(* IEC 61131-3 sources: Summary-ETFA22/ahorn/test/benchmark/dissertation/PPU/ST (part 5) *)

        //End of: edu.kit.iti.formal.automation.st.IntroduceStateEnumVariable

        //Running pipeline step: edu.kit.iti.formal.automation.st.TranslationSfcToStOld$IntroduceTransitVariable

        //End of: edu.kit.iti.formal.automation.st.TranslationSfcToStOld$IntroduceTransitVariable

        //Running pipeline step: edu.kit.iti.formal.automation.st.TranslationSfcToStOld$TheBigStateCase

        CASE _state OF
            STATES_STAMP#Init:
                __transit := FALSE;
                IF TRUE THEN
                    __transit := TRUE;
                    _state := STATES_STAMP#Start_Stamp;
                END_IF

            STATES_STAMP#Start_Stamp:
                __transit := FALSE;
                Start_Stamp_active();
                IF interconnectStampStartCommand THEN
                    __transit := TRUE;
                    _state := STATES_STAMP#Green_Lamp;
                END_IF

            STATES_STAMP#Green_Lamp:
                __transit := FALSE;
                Green_Lamp_active();
                IF TRUE THEN
                    __transit := TRUE;
                    _state := STATES_STAMP#Stamp_Init_1;
                END_IF

            STATES_STAMP#Stamp_Init_1:
                __transit := FALSE;
                Stamp_Init_1_active();
                IF StampSliderSensorMovedIn THEN
                    __transit := TRUE;
                    _state := STATES_STAMP#Stamp_Init_2;
                END_IF

            STATES_STAMP#Stamp_Init_2:
                __transit := FALSE;
                Stamp_Init_2_active();
                IF StampSliderSensorMovedOut THEN
                    __transit := TRUE;
                    _state := STATES_STAMP#Stamp_Init_3;
                END_IF

            STATES_STAMP#Stamp_Init_3:
                __transit := FALSE;
                Stamp_Init_3_active();
                IF StampLowered THEN
                    __transit := TRUE;
                    _state := STATES_STAMP#Stamp_Init_4;
                END_IF

            STATES_STAMP#Stamp_Init_4:
                __transit := FALSE;
                Stamp_Init_4_active();
                IF StampUp THEN
                    __transit := TRUE;
                    _state := STATES_STAMP#Interstep;
                END_IF

            STATES_STAMP#Interstep:
                __transit := FALSE;
                Interstep_active();
                IF StartVar THEN
                    __transit := TRUE;
                    _state := STATES_STAMP#Intertsep_2;
                END_IF

            STATES_STAMP#Intertsep_2:
                __transit := FALSE;
                IF StampSliderFilled THEN
                    __transit := TRUE;
                    _state := STATES_STAMP#Step0;
                END_IF

            STATES_STAMP#Step0:
                __transit := FALSE;
                IF CraneUp THEN
                    __transit := TRUE;
                    _state := STATES_STAMP#StampSliderBack;
                END_IF

            STATES_STAMP#StampSliderBack:
                __transit := FALSE;
                StampSliderBack_active();
                IF StampSliderSensorMovedIn THEN
                    __transit := TRUE;
                    _state := STATES_STAMP#StampProcess;
                END_IF

            STATES_STAMP#StampProcess:
                __transit := FALSE;
                StampProcess_active();
                IF StampLowered THEN
                    __transit := TRUE;
                    _state := STATES_STAMP#Step1;
                END_IF

            STATES_STAMP#Step1:
                __transit := FALSE;
                Step1_active();
                IF interconnect THEN
                    __transit := TRUE;
                    _state := STATES_STAMP#StampSliderForward;
                END_IF

            STATES_STAMP#StampSliderForward:
                __transit := FALSE;
                StampSliderForward_active();
                IF StampSliderMovedOut THEN
                    __transit := TRUE;
                    _state := STATES_STAMP#Step2;
                END_IF

            STATES_STAMP#Step2:
                __transit := FALSE;
                IF (((AnalogCranePosition > 16160) AND (AnalogCranePosition < 16260)) AND NOT StampSliderFilled) THEN
                    __transit := TRUE;
                    _state := STATES_STAMP#Interstep;
                END_IF

                    END_CASE
        //End of: edu.kit.iti.formal.automation.st.TranslationSfcToStOld$TheBigStateCase

        //Running pipeline step: edu.kit.iti.formal.automation.st.SfcFlagIntroduction

    END_IF
    //End of: edu.kit.iti.formal.automation.st.SfcFlagIntroduction

END_FUNCTION_BLOCK

PROGRAM Main
    VAR_OUTPUT
        Actuator_AnalogCranePressure : INT := INT#0;
        Actuator_CraneLower : BOOL := FALSE;
        Actuator_CraneTurnClockwise : BOOL := FALSE;
        Actuator_CraneTurnCounterclockwise : BOOL := FALSE;
        Actuator_MagazinGreenLamp : BOOL := FALSE;
        Actuator_MagazinSlider : BOOL := FALSE;
        Actuator_MagazinVacuumOff : BOOL := FALSE;
        Actuator_MagazinVacuumOn : BOOL := FALSE;
        Actuator_MagazinWhiteLamp : BOOL := FALSE;
        Actuator_PusherY1 : BOOL := FALSE;
        Actuator_PusherY2 : BOOL := FALSE;
        Actuator_SorterConveyorTowardsCrane : BOOL := FALSE;
        Actuator_SorterConveyorTowardsStacker : BOOL := FALSE;
        Actuator_SorterGreenLampConveyor : BOOL := FALSE;
        Actuator_SorterWhiteLampConveyor : BOOL := FALSE;
        Actuator_StampGreenLamp : BOOL := FALSE;
        Actuator_StampPusher : BOOL := FALSE;
        Actuator_StampSliderMovedIn : BOOL := FALSE;
        Actuator_StampSliderMovedOut : BOOL := FALSE;
        Actuator_StampWhiteLamp : BOOL := FALSE;
    END_VAR

    VAR
        Conveyor : Conveyor := (SFCReset:=FALSE, Timer_Conveyor_Runtime:=(Q:=FALSE, PT:=UINT#0, IN:=FALSE, ET:=UINT#0), SorterStartButton:=FALSE, interconnect_Conveyor_Test:=FALSE, SorterConveyorTowardsCrane:=FALSE, interconnectConveyorStartCommand:=FALSE, SFCInit:=FALSE, interconnectConveyorTerminationCommand:=FALSE, SorterConveyorTowardsStacker:=FALSE, interconnect_Conveyor_Runtime:=FALSE, Timer_Conveyor_Test:=(Q:=FALSE, PT:=UINT#0, IN:=FALSE, ET:=UINT#0), SorterLightbarrierCraneInterface:=FALSE, SorterSwitchManuellAutomatic:=FALSE, StartVar:=FALSE, SorterGreenLampConveyor:=FALSE, StartCommandConveyor:=FALSE, Duration_Conveyor_Test:=TIME#1000.0ms, Duration_Conveyor_Runtime:=TIME#4500.0ms, SorterWhiteLampConveyor:=FALSE);
        Crane : Crane := (SliderMovedOut:=FALSE, CraneTurnCounterclockwise:=FALSE, WorkpieceReady:=FALSE, StampLowered:=FALSE, Duration1:=TIME#1500.0ms, StampSliderSensorMovedOut:=FALSE, TimeDelay_Timer_interconnect:=FALSE, MagazinOpticalSensor:=FALSE, StartVar:=FALSE, StartButtonMagazin:=FALSE, actualtime1:=TIME#, AnalogCranePressure:=INT#0, SFCReset:=FALSE, AnalogCranePosition:=INT#0, MagazinVacuumOff:=FALSE, CraneSucked:=FALSE, MagazinSlider:=FALSE, MagazinVacuumOn:=FALSE, interconnectCraneStartCommand:=FALSE, SFCInit:=FALSE, StartCommandCrane:=FALSE, TimeDelay_Timer_Duration:=TIME#50.0ms, interconnect:=FALSE, StampSliderFilled:=FALSE, CraneTurnClockwise:=FALSE, CraneUp:=FALSE, MagazinCapacitiveSensor:=FALSE, CraneLower:=FALSE, SliderNotMovedOut:=FALSE, CraneDown:=FALSE, TimeDelay_Timer:=(Q:=FALSE, PT:=UINT#0, IN:=FALSE, ET:=UINT#0), Timer1:=(Q:=FALSE, PT:=UINT#0, IN:=FALSE, ET:=UINT#0));
        Mag : Magazin := (SliderMovedOut:=FALSE, MagazinGreenLamp:=FALSE, interconnectMagazinStartCommand:=FALSE, SFCReset:=FALSE, AnalogCranePosition:=INT#0, CraneTurnCounterclockwise:=FALSE, MagazinVacuumOff:=FALSE, WorkpieceReady:=FALSE, CraneSucked:=FALSE, MagazinSlider:=FALSE, MagazinVacuumOn:=FALSE, MagazinWhiteLamp:=FALSE, SFCInit:=FALSE, StartCommandMagazin:=FALSE, CraneOnConveyor:=FALSE, CraneTurnClockwise:=FALSE, CraneUp:=FALSE, StartVar:=FALSE, CraneLower:=FALSE, SliderNotMovedOut:=FALSE, StartButtonMagazin:=FALSE, CraneOnMagazin:=FALSE, CraneDown:=FALSE);
        Pusher : Pusher := (Slide2_metal:=INT#1, Timer_Slide2_White:=(Q:=FALSE, PT:=UINT#0, IN:=FALSE, ET:=UINT#0), SorterPusher1MovedIn:=FALSE, SorterPusher2MovedIn:=FALSE, Slide3_white:=INT#1, Slide3_black:=INT#1, Timer_Slide1_Black:=(Q:=FALSE, PT:=UINT#0, IN:=FALSE, ET:=UINT#0), PusherY2:=FALSE, Priority_Var_Metal:=INT#3, PusherY1:=FALSE, SFCReset:=FALSE, SorterCapacitiveSensorPusher2:=FALSE, SorterCapacitiveSensorPusher1:=FALSE, Timer_Slide1_White:=(Q:=FALSE, PT:=UINT#0, IN:=FALSE, ET:=UINT#0), Timer_Slide2_Metal:=(Q:=FALSE, PT:=UINT#0, IN:=FALSE, ET:=UINT#0), Slide3_metal:=INT#1, Duration_Slide1_Metal:=TIME#300.0ms, Duration_Slide1_Black:=TIME#950.0ms, interconnect_Slide1_White:=FALSE, interconnect_Slide2_Metal:=FALSE, SorterPusher2MovedOut:=FALSE, Slide2_white:=INT#1, Priority_Var_Black:=INT#3, Duration_Slide2_Black:=TIME#2000.0ms, SorterLightnessSensorPusher2:=FALSE, SorterPusher1MovedOut:=FALSE, SorterStartButton:=FALSE, SorterLightnessSensorPusher1:=FALSE, Duration3:=TIME#200.0ms, Duration2:=TIME#2000.0ms, Slide1_black:=INT#1, interconnect_Slide2_White:=FALSE, SorterLightbarrierCraneInterface:=FALSE, StartVar:=FALSE, Duration_Slide2_White:=TIME#370.0ms, interconnect_Slide2_Black:=FALSE, SorterLightnessSensorPusher3:=FALSE, Slide1_white:=INT#1, interconnect3:=FALSE, interconnect2:=FALSE, interconnect_Slide1_Metal:=FALSE, Slide1_metal:=INT#1, SFCInit:=FALSE, Priority_Var_White:=INT#3, Slide2_black:=INT#1, Duration_Slide2_Metal:=TIME#370.0ms, interconnect_Slide1_Black:=FALSE, SorterLightnesssensorCraneInterfaceInverse:=FALSE, Timer_Slide1_Metal:=(Q:=FALSE, PT:=UINT#0, IN:=FALSE, ET:=UINT#0), Timer2:=(Q:=FALSE, PT:=UINT#0, IN:=FALSE, ET:=UINT#0), Timer_Slide2_Black:=(Q:=FALSE, PT:=UINT#0, IN:=FALSE, ET:=UINT#0), Duration_Slide1_White:=TIME#300.0ms, Timer3:=(Q:=FALSE, PT:=UINT#0, IN:=FALSE, ET:=UINT#0));
        Stamp : Stamp := (StampLowered:=FALSE, StampSliderSensorMovedOut:=FALSE, interconnectStampStartCommand:=FALSE, CraneOnConveyor:=FALSE, CranePositionStamp:=FALSE, StampSliderMovedOut:=FALSE, StartVar:=FALSE, StampPusher:=FALSE, StampWhiteLamp:=FALSE, StampPressure:=FALSE, SFCReset:=FALSE, StampGreenLamp:=FALSE, AnalogCranePosition:=INT#0, CraneSucked:=FALSE, Duration:=TIME#500.0ms, SFCInit:=FALSE, StampStartButton:=FALSE, StampSliderSensorMovedIn:=FALSE, interconnect:=FALSE, StampSliderFilled:=FALSE, CraneUp:=FALSE, StampSliderMovedIn:=FALSE, Timer:=(Q:=FALSE, PT:=UINT#0, IN:=FALSE, ET:=UINT#0), StartCommandStamp:=FALSE, CraneDown:=FALSE, StampUp:=FALSE);
    END_VAR

    VAR_INPUT
        Sensor_AnalogCranePosition : INT := INT#0;
        Sensor_CraneDown : BOOL := FALSE;
        Sensor_CraneOnConveyor : BOOL := FALSE;
        Sensor_CraneOnMagazin : BOOL := FALSE;
        Sensor_CranePosition : BOOL := FALSE;
        Sensor_CranePositionStamp : BOOL := FALSE;
        Sensor_CraneSucked : BOOL := FALSE;
        Sensor_CraneUp : BOOL := FALSE;
        Sensor_MagazinCapacitiveSensor : BOOL := FALSE;
        Sensor_MagazinEmergencyStop : BOOL := FALSE;
        Sensor_MagazinOpticalSensor : BOOL := FALSE;
        Sensor_MagazinSwitchManuellAutomatic : BOOL := FALSE;
        Sensor_SliderMovedOut : BOOL := FALSE;
        Sensor_SliderNotMovedOut : BOOL := FALSE;
        Sensor_SorterCapacitiveSensorPusher1 : BOOL := FALSE;
        Sensor_SorterCapacitiveSensorPusher2 : BOOL := FALSE;
        Sensor_SorterEmergencyStop : BOOL := FALSE;
        Sensor_SorterLightbarrierCraneInterface : BOOL := FALSE;
        Sensor_SorterLightnessSensorPusher1 : BOOL := FALSE;
        Sensor_SorterLightnessSensorPusher2 : BOOL := FALSE;
        Sensor_SorterLightnessSensorPusher3 : BOOL := FALSE;
        Sensor_SorterLightnesssensorCraneInterfaceInverse : BOOL := FALSE;
        Sensor_SorterPusher1MovedIn : BOOL := FALSE;
        Sensor_SorterPusher1MovedOut : BOOL := FALSE;
        Sensor_SorterPusher2MovedIn : BOOL := FALSE;
        Sensor_SorterPusher2MovedOut : BOOL := FALSE;
        Sensor_SorterStartButton : BOOL := FALSE;
        Sensor_SorterSwitchManuellAutomatic : BOOL := FALSE;
        Sensor_StampEmergencyStop : BOOL := FALSE;
        Sensor_StampLowered : BOOL := FALSE;
        Sensor_StampSliderFilled : BOOL := FALSE;
        Sensor_StampSliderSensorMovedIn : BOOL := FALSE;
        Sensor_StampSliderSensorMovedOut : BOOL := FALSE;
        Sensor_StampStartButton : BOOL := FALSE;
        Sensor_StampSwitchManuellAutomatic : BOOL := FALSE;
        Sensor_StampUp : BOOL := FALSE;
        Sensor_StartButtonMagazin : BOOL := FALSE;
        Sensor_WorkpieceReady : BOOL := FALSE;
    END_VAR

    Mag.SliderNotMovedOut := Sensor_SliderNotMovedOut;
    Mag.SliderMovedOut := Sensor_SliderMovedOut;
    Mag.CraneOnMagazin := Sensor_CraneOnMagazin;
    Mag.CraneDown := Sensor_CraneDown;
    Mag.CraneUp := Sensor_CraneUp;
    Mag.CraneOnConveyor := Sensor_CraneOnConveyor;
    Mag.WorkpieceReady := Sensor_WorkpieceReady;
    Mag.AnalogCranePosition := Sensor_AnalogCranePosition;
    Mag.StartButtonMagazin := Sensor_StartButtonMagazin;
    Actuator_MagazinSlider := Mag.MagazinSlider;
    Actuator_MagazinGreenLamp := Mag.MagazinGreenLamp;
    Crane.CraneUp := Sensor_CraneUp;
    Crane.CraneDown := Sensor_CraneDown;
    Crane.CraneSucked := Sensor_CraneSucked;
    Crane.MagazinCapacitiveSensor := Sensor_MagazinCapacitiveSensor;
    Crane.SliderMovedOut := Sensor_SliderMovedOut;
    Crane.WorkpieceReady := Sensor_WorkpieceReady;
    Crane.MagazinOpticalSensor := Sensor_MagazinOpticalSensor;
    Crane.StampSliderFilled := Sensor_StampSliderFilled;
    Crane.StampSliderSensorMovedOut := Sensor_StampSliderSensorMovedOut;
    Crane.StampLowered := Sensor_StampLowered;
    Crane.AnalogCranePosition := Sensor_AnalogCranePosition;
    Crane.StartButtonMagazin := Sensor_StartButtonMagazin;
    Actuator_CraneTurnCounterclockwise := Crane.CraneTurnCounterclockwise;
    Actuator_CraneTurnClockwise := Crane.CraneTurnClockwise;
    Actuator_CraneLower := Crane.CraneLower;
    Actuator_MagazinVacuumOff := Crane.MagazinVacuumOff;
    Actuator_MagazinVacuumOn := Crane.MagazinVacuumOn;
    Actuator_AnalogCranePressure := Crane.AnalogCranePressure;
    Stamp.StampSliderSensorMovedOut := Sensor_StampSliderSensorMovedOut;
    Stamp.StampSliderSensorMovedIn := Sensor_StampSliderSensorMovedIn;
    Stamp.StampSliderFilled := Sensor_StampSliderFilled;
    Stamp.StampUp := Sensor_StampUp;
    Stamp.StampLowered := Sensor_StampLowered;
    Stamp.CraneDown := Sensor_CraneDown;
    Stamp.CraneUp := Sensor_CraneUp;
    Stamp.CraneSucked := Sensor_CraneSucked;
    Stamp.CranePositionStamp := Sensor_CranePositionStamp;
    Stamp.CraneOnConveyor := Sensor_CraneOnConveyor;
    Stamp.AnalogCranePosition := Sensor_AnalogCranePosition;
    Stamp.StampStartButton := Sensor_StampStartButton;
    Actuator_StampSliderMovedOut := Stamp.StampSliderMovedOut;
    Actuator_StampSliderMovedIn := Stamp.StampSliderMovedIn;
    Actuator_StampWhiteLamp := Stamp.StampWhiteLamp;
    Actuator_StampPusher := Stamp.StampPusher;
    Actuator_StampGreenLamp := Stamp.StampGreenLamp;
    Conveyor.SorterStartButton := Sensor_SorterStartButton;
    Conveyor.SorterSwitchManuellAutomatic := Sensor_SorterSwitchManuellAutomatic;
    Conveyor.SorterLightbarrierCraneInterface := Sensor_SorterLightbarrierCraneInterface;
    Actuator_SorterConveyorTowardsStacker := Conveyor.SorterConveyorTowardsStacker;
    Actuator_SorterConveyorTowardsCrane := Conveyor.SorterConveyorTowardsCrane;
    Actuator_SorterGreenLampConveyor := Conveyor.SorterGreenLampConveyor;
    Actuator_SorterWhiteLampConveyor := Conveyor.SorterWhiteLampConveyor;
    Pusher.SorterLightnesssensorCraneInterfaceInverse := Sensor_SorterLightnesssensorCraneInterfaceInverse;
    Pusher.SorterLightbarrierCraneInterface := Sensor_SorterLightbarrierCraneInterface;
    Pusher.SorterCapacitiveSensorPusher1 := Sensor_SorterCapacitiveSensorPusher1;
    Pusher.SorterLightnessSensorPusher1 := Sensor_SorterLightnessSensorPusher1;
    Pusher.SorterCapacitiveSensorPusher2 := Sensor_SorterCapacitiveSensorPusher2;
    Pusher.SorterLightnessSensorPusher2 := Sensor_SorterLightnessSensorPusher2;
    Pusher.SorterLightnessSensorPusher3 := Sensor_SorterLightnessSensorPusher3;
    Pusher.SorterPusher1MovedOut := Sensor_SorterPusher1MovedOut;
    Pusher.SorterPusher1MovedIn := Sensor_SorterPusher1MovedIn;
    Pusher.SorterPusher2MovedOut := Sensor_SorterPusher2MovedOut;
    Pusher.SorterPusher2MovedIn := Sensor_SorterPusher2MovedIn;
    Pusher.SorterStartButton := Sensor_SorterStartButton;
    Actuator_PusherY1 := Pusher.PusherY1;
    Actuator_PusherY2 := Pusher.PusherY2;
    IF ((Sensor_SorterEmergencyStop AND Sensor_StampEmergencyStop) AND Sensor_MagazinEmergencyStop) THEN
        Mag();
        Crane();
        Stamp();
        Conveyor();
        Pusher();
        IF ((Actuator_SorterGreenLampConveyor AND Actuator_MagazinGreenLamp) AND Actuator_StampGreenLamp) THEN
            IF (((Stamp.StartCommandStamp AND Crane.StartCommandCrane) AND Conveyor.StartCommandConveyor) AND Mag.StartCommandMagazin) THEN
                Crane.StartVar := TRUE;
                Conveyor.StartVar := TRUE;
                Mag.StartVar := TRUE;
                Pusher.StartVar := TRUE;
                Stamp.StartVar := TRUE;
            END_IF
        END_IF
        Crane.SFCReset := FALSE;
        Conveyor.SFCReset := FALSE;
        Mag.SFCReset := FALSE;
        Pusher.SFCReset := FALSE;
        Stamp.SFCReset := FALSE;
    ELSIF ((NOT Sensor_SorterEmergencyStop OR NOT Sensor_StampEmergencyStop) OR NOT Sensor_MagazinEmergencyStop) THEN
        Actuator_MagazinSlider := FALSE;
        Actuator_CraneLower := FALSE;
        Actuator_MagazinVacuumOn := FALSE;
        Actuator_MagazinVacuumOff := TRUE;
        Actuator_MagazinGreenLamp := FALSE;
        Actuator_CraneTurnCounterclockwise := FALSE;
        Actuator_CraneTurnClockwise := FALSE;
        Actuator_SorterConveyorTowardsStacker := FALSE;
        Actuator_SorterConveyorTowardsCrane := FALSE;
        Actuator_SorterGreenLampConveyor := FALSE;
        Actuator_PusherY1 := FALSE;
        Actuator_PusherY2 := FALSE;
        Actuator_StampSliderMovedOut := TRUE;
        Actuator_StampSliderMovedIn := FALSE;
        Actuator_StampGreenLamp := FALSE;
        Actuator_StampPusher := FALSE;
        Actuator_AnalogCranePressure := INT#0;
        Crane.SFCReset := TRUE;
        Conveyor.SFCReset := TRUE;
        Mag.SFCReset := TRUE;
        Pusher.SFCReset := TRUE;
        Stamp.SFCReset := TRUE;
        Crane.StartVar := FALSE;
        Conveyor.StartVar := FALSE;
        Mag.StartVar := FALSE;
        Pusher.StartVar := FALSE;
        Stamp.StartVar := FALSE;
    END_IF
END_PROGRAM
FUNCTION_BLOCK CTD

    VAR_INPUT
        CD : BOOL := FALSE;
        LD : BOOL := FALSE;
        PV : INT := INT#0;
    END_VAR

    VAR_OUTPUT
        CV : INT := INT#0;
        Q : BOOL := FALSE;
    END_VAR

    IF LD THEN
        CV := PV;
    ELSIF (CU AND (CV > INT#0)) THEN
        CV := (CV - INT#1);
    END_IF
    Q := (CV <= INT#0);
END_FUNCTION_BLOCK

FUNCTION_BLOCK CTU

    VAR_INPUT
        CU : BOOL := FALSE;
        PV : INT := INT#0;
        R : BOOL := FALSE;
    END_VAR

    VAR_OUTPUT
        CV : INT := INT#0;
        Q : BOOL := FALSE;
    END_VAR

    IF R THEN
        CV := INT#0;
    ELSIF (CU AND (CV < PV)) THEN
        CV := (CV + INT#1);
    END_IF
    Q := (CV >= PV);
END_FUNCTION_BLOCK

FUNCTION_BLOCK R_TRIG

    VAR_INPUT
        CLK : BOOL := FALSE;
    END_VAR

    VAR
        M : BOOL := FALSE;
    END_VAR

    VAR_OUTPUT
        Q : BOOL := FALSE;
    END_VAR

    Q := (CLK AND NOT M);
    M := CLK;
END_FUNCTION_BLOCK

FUNCTION_BLOCK F_TRIG

    VAR_INPUT
        CLK : BOOL := FALSE;
    END_VAR

    VAR
        M : BOOL := TRUE;
    END_VAR

    VAR_OUTPUT
        Q : BOOL := FALSE;
    END_VAR

    Q := (NOT CLK AND NOT M);
    M := NOT CLK;
END_FUNCTION_BLOCK

FUNCTION SEL : ANY

    VAR_INPUT
        G : BOOL := FALSE;
        a : ANY;
        b : ANY;
    END_VAR

    VAR_OUTPUT
        SEL : ANY;
    END_VAR

    IF G THEN
        SEL := a;
    ELSE
        SEL := b;
    END_IF
END_FUNCTION

FUNCTION MAX : ANY_INT

    VAR_OUTPUT
        MAX : ANY_INT;
    END_VAR

    VAR_INPUT
        in0 : ANY_INT;
        in1 : ANY_INT;
    END_VAR

    MAX := sel((in0 >= in1), in0, in1);
END_FUNCTION

FUNCTION MIN : ANY_INT

    VAR_OUTPUT
        MIN : ANY_INT;
    END_VAR

    VAR_INPUT
        in0 : ANY_INT;
        in1 : ANY_INT;
    END_VAR

    MIN := sel((in0 <= in1), in0, in1);
END_FUNCTION

FUNCTION LIMIT : INT

    VAR_OUTPUT
        LIMIT : INT := INT#0;
    END_VAR

    VAR_INPUT
        in : ANY_INT;
        max : ANY_INT;
        min : ANY_INT;
    END_VAR

    LIMIT := MAX(min, MIN(in, max));
END_FUNCTION

FUNCTION ERROR : ANY

    VAR_OUTPUT
        ERROR : ANY;
    END_VAR

    VAR
        msg : STRING := WSTRING#"";
    END_VAR

END_FUNCTION

FUNCTION SMV : ANY

    VAR_OUTPUT
        SMV : ANY;
    END_VAR

    VAR_INPUT
        code : STRING := WSTRING#"";
    END_VAR

END_FUNCTION

FUNCTION_BLOCK TON

    VAR_OUTPUT
        ET : UINT := UINT#0;
        Q : BOOL := FALSE;
    END_VAR

    VAR_INPUT
        IN : BOOL := FALSE;
        PT : UINT := UINT#0;
    END_VAR

    IF IN THEN
        Q := (ET = UINT#0);
        IF (ET > UINT#0) THEN
            ET := (ET - UINT#1);
        ELSE
            ET := UINT#0;
        END_IF
    ELSE
        Q := FALSE;
        ET := PT;
    END_IF
END_FUNCTION_BLOCK

TYPE SFC_STEPS: STRUCT

        T :TIME
        X :BOOL
        _T :TIME
        _X :BOOLEND_STRUCT;

END_TYPE

TYPE
    STATES_CONVEYOR : (Init, Start_Conveyor, Green_Lamp, Conveyor_Init, Conveyor_init_2, Interstep, Step0, Conveyor_Towards_Stacker, Runtime_Conveyor, Conveyor_pause, Conveyor_Stop_Empty_Magazin);
    STATES_CRANE : (Init, Start_Crane, Crane_Init, Crane_Init_2, Interstep, Interstep_2, TimeDelay, Interstep_3, Turn_Right, Magazin_Stop, Crane_Lower, Step0, Crane_Lift_Magazin, Crane_Turn_Left_NOT_Metallic, Crane_On_Conveyor, Stamp_Pressure_Profile_Set_Metallic, Crane_Lift_Magazin_Metallic, Crane_Turn_Left_Metallic, Crane_On_Stamp_Metallic, release_Workpiece, Crane_Go_Up, Stamp_Pressure_Profile_Set_White, Crane_Lift_Magazin_White, Crane_Turn_Left_White, Crane_On_Stamp_White, release_Workpiece_White, Crane_Go_Up_White, Step3, Step2, pause, Turn_Right_Black, Magazin_Stop_Black, Crane_Lift_NOT_Metallic_Black, Crane_Turn_Left_NOT_Metallic_Black, Crane_On_Conveyor_Not_Metallica_Black, release_Black, Crane_Lift_Conveyor_Black, Crane_Turn_Left_Back_To_Stamp, Crane_On_Stamp_Stop_Black, Step4, Reset_interconnect, Lower_Crane, Suck_At_Stamp, Crane_Lift_At_Stamp, Crane_Turn_Left_From_Stamp, Crane_On_Conveyor_Metallic, release, Crane_Lift_Conveyor, No_Workpiece_ready, Crane_Turn_Left_Metallic2, Crane_On_Stamp_Metallic2, Interstep_4, Crane_On_Stamp_Metallic2_Lower, Suck_At_Stamp2, Crane_Lift_At_Stamp2, Crane_Turn_Right_From_Stamp, Crane_On_Conveyor_Metallic2, release2, Crane_Lift_Conveyor2, Turn_Right_Final, Magazin_Stop_Final);
    STATES_MAGAZIN : (Init, Start_Magazin, Green_Lamp, Magazin_Init, Magazin_Init_2, Interstep, convey, Step0, Slider_Move_Back, Step1);
    STATES_PUSHER : (Init, Interstep, Interstep_2, Check_For_Black, Third_Slide_black_workpieces, Wait_Black, Reset_interconnect3, Second_Slide_black_workpieces, Second_Slide_Timer_Black, PusherY2_Move_Out_Black, Wait_Y2_Black, PusherY2_Move_In_Black, Reset_interconnect_Slide2_Black, First_Slide_black_workpieces, First_Slide_Timer_Black, PusherY1_Move_Out_Black, Wait_Y1_Black, PusherY1_Move_In_Black, Reset_interconnect_Slide1_Black, Check_For_White, First_Slide_white_workpieces, First_Slide_Timer_White, PusherY1_Move_Out_White, Wait_Y1_White, PusherY1_Move_In_White, Reset_interconnect_Slide1_White, Second_Slide_white_workpieces, Second_Test_For_White, Second_Slide_Timer_White, PusherY2_Move_Out_White, Wait_Y2_White, PusherY2_Move_In_White, Reset_interconnect_Slide2_White, Third_Slide_white_workpieces, Wait_White, Reset_interconnect_Slide3_White, Check_For_Metal, First_Slide_metal_workpieces, First_Slide_Timer_Metal, PusherY1_Move_Out_Metal, Wait_Y1_Metal, PusherY1_Move_In_Metal, Reset_interconnect_Slide1_Metal, Second_Slide_metal_workpieces, Second_Test_For_Metal, Second_Slide_Timer_Metal, PusherY2_Move_Out_Metal, Wait_Y2_Metal, PusherY2_Move_In_Metal, Reset_interconnect_Slide2_Metal, Third_Slide_metal_workpieces, Wait_Metal, Reset_interconnect_Slide3_Metal);
    STATES_STAMP : (Init, Start_Stamp, Green_Lamp, Stamp_Init_1, Stamp_Init_2, Stamp_Init_3, Stamp_Init_4, Interstep, Intertsep_2, Step0, StampSliderBack, StampProcess, Step1, StampSliderForward, Step2);
END_TYPE

(* ---- Scenario1_Final.st ---- *)
TYPE
    CraneStates : (CraneSFCInit, StartCrane, CraneInit, CraneInit2, Interstep, Interstep2, TimeDelay, TurnRight,
                   InterstepCheckWorkpiece, StackStop, CraneLiftStack, CraneTurnLeft, CraneOnConveyorState,
                   release, CraneLiftConveyor, CraneStop);
    StackStates : (StackSFCInit, StartStack, GreenLamp, StackInit, StackInit2, Interstep, convey, Step0,
                   SliderMoveBack, Step1);
END_TYPE

FUNCTION_BLOCK Crane
VAR_INPUT
    CraneDown : BOOL := FALSE;
    CraneOnConveyor : BOOL := FALSE;
    CraneOnStack : BOOL := FALSE;
    CraneSucked : BOOL := FALSE;
    CraneUp : BOOL := FALSE;
    SFCReset : BOOL := FALSE;
    SliderMovedOut : BOOL := FALSE;
    SliderNotMovedOut : BOOL := FALSE;
    StartButtonStack : BOOL := FALSE;
    StartVar : BOOL := FALSE;
    WorkpieceReady : BOOL := FALSE;
END_VAR
VAR
    SFCInit : BOOL := FALSE;
    SFCPause : BOOL := FALSE;
    CraneState : CraneStates := CraneStates#CraneSFCInit;
    Timer : TON;
    TimerDuration : TIME := TIME#50.0ms;
    Timerinterconnect : BOOL := FALSE;
    interconnectCraneStartCommand : BOOL := FALSE;
END_VAR
VAR_OUTPUT
    CraneLower : BOOL := FALSE;
    CraneTurnClockwise : BOOL := FALSE;
    CraneTurnCounterClockwise : BOOL := FALSE;
    StackVacuumOff : BOOL := FALSE;
    StackVacuumOn : BOOL := FALSE;
    StartCommandCrane : BOOL := FALSE;
END_VAR

IF (SFCInit OR SFCReset) THEN
    CraneDown := FALSE;
    CraneLower := FALSE;
    CraneOnConveyor := FALSE;
    CraneOnStack := FALSE;
    CraneSucked := FALSE;
    CraneTurnClockwise := FALSE;
    CraneTurnCounterClockwise := FALSE;
    CraneUp := FALSE;
    StackVacuumOff := FALSE;
    StackVacuumOn := FALSE;
    SFCInit := FALSE;
    SFCReset := FALSE;
    SliderMovedOut := FALSE;
    SliderNotMovedOut := FALSE;
    StartButtonStack := FALSE;
    StartCommandCrane := FALSE;
    StartVar := FALSE;
    Timer.ET := INT#0;
    Timer.IN := FALSE;
    Timer.PT := INT#0;
    Timer.Q := FALSE;
    TimerDuration := TIME#50ms;
    Timerinterconnect := FALSE;
    WorkpieceReady := FALSE;
    CraneState := CraneStates#CraneSFCInit;
    interconnectCraneStartCommand := FALSE;
END_IF;

IF NOT (SFCInit OR SFCPause) THEN
    CASE CraneState OF
        CraneStates#CraneSFCInit:
            IF TRUE THEN
                CraneState := CraneStates#StartCrane;
            END_IF;

        CraneStates#StartCrane:
            CraneLower := FALSE;
            StackVacuumOff := TRUE;
            StackVacuumOn := FALSE;
            CraneTurnCounterClockwise := FALSE;
            CraneTurnClockwise := FALSE;
            StartVar := FALSE;
            StartCommandCrane := FALSE;
            IF (StartButtonStack = TRUE) THEN
                interconnectCraneStartCommand := TRUE;
            END_IF;
            IF interconnectCraneStartCommand THEN
                CraneState := CraneStates#CraneInit;
            END_IF;

        CraneStates#CraneInit:
            CraneLower := TRUE;
            interconnectCraneStartCommand := FALSE;
            IF CraneDown THEN
                CraneState := CraneStates#CraneInit2;
            END_IF;

        CraneStates#CraneInit2:
            CraneLower := FALSE;
            IF CraneUp THEN
                CraneState := CraneStates#Interstep;
            END_IF;

        CraneStates#Interstep:
            StartCommandCrane := TRUE;
            IF StartVar THEN
                CraneState := CraneStates#Interstep2;
            END_IF;

        CraneStates#Interstep2:
            IF SliderMovedOut THEN
                CraneState := CraneStates#TimeDelay;
            END_IF;

        CraneStates#TimeDelay:
            Timer(IN := TRUE, PT := TimerDuration);
            Timerinterconnect := Timer.Q;
            IF Timerinterconnect THEN
                CraneState := CraneStates#TurnRight;
            END_IF;

        CraneStates#TurnRight:
            CraneTurnClockwise := TRUE;
            CraneTurnCounterClockwise := FALSE;
            IF CraneOnStack THEN
                CraneState := CraneStates#InterstepCheckWorkpiece;
            END_IF;

        CraneStates#InterstepCheckWorkpiece:
            IF WorkpieceReady THEN
                CraneState := CraneStates#StackStop;
            ELSIF NOT WorkpieceReady THEN
                CraneState := CraneStates#CraneStop;
            END_IF;

        CraneStates#StackStop:
            CraneTurnClockwise := FALSE;
            CraneTurnCounterClockwise := FALSE;
            StackVacuumOn := TRUE;
            StackVacuumOff := FALSE;
            CraneLower := TRUE;
            IF CraneSucked THEN
                CraneState := CraneStates#CraneLiftStack;
            END_IF;

        CraneStates#CraneLiftStack:
            CraneLower := FALSE;
            IF CraneUp THEN
                CraneState := CraneStates#CraneTurnLeft;
            END_IF;

        CraneStates#CraneTurnLeft:
            CraneTurnCounterClockwise := TRUE;
            CraneTurnClockwise := FALSE;
            IF CraneOnConveyor THEN
                CraneState := CraneStates#CraneOnConveyorState;
            END_IF;

        CraneStates#CraneOnConveyorState:
            CraneTurnCounterClockwise := FALSE;
            CraneTurnClockwise := FALSE;
            CraneLower := TRUE;
            IF CraneDown THEN
                CraneState := CraneStates#release;
            END_IF;

        CraneStates#release:
            StackVacuumOff := TRUE;
            StackVacuumOn := FALSE;
            IF TRUE THEN
                CraneState := CraneStates#CraneLiftConveyor;
            END_IF;

        CraneStates#CraneLiftConveyor:
            CraneLower := FALSE;
            IF TRUE THEN
                CraneState := CraneStates#Interstep;
            END_IF;

        CraneStates#CraneStop:
            IF TRUE THEN
                CraneState := CraneStates#StartCrane;
            END_IF;
    END_CASE;
END_IF;
END_FUNCTION_BLOCK

FUNCTION_BLOCK Stack
VAR_INPUT
    CraneDown : BOOL := FALSE;
    CraneOnConveyor : BOOL := FALSE;
    CraneOnStack : BOOL := FALSE;
    CraneSucked : BOOL := FALSE;
    CraneUp : BOOL := FALSE;
    SFCReset : BOOL := FALSE;
    SliderMovedOut : BOOL := FALSE;
    SliderNotMovedOut : BOOL := FALSE;
    StartButtonStack : BOOL := FALSE;
    StartVar : BOOL := FALSE;
    WorkpieceReady : BOOL := FALSE;
END_VAR
VAR
    SFCInit : BOOL := FALSE;
    SFCPause : BOOL := FALSE;
    StackState : StackStates := StackStates#StackSFCInit;
    interconnectStackStartCommand : BOOL := FALSE;
END_VAR
VAR_OUTPUT
    StackGreenLamp : BOOL := FALSE;
    StackSlider : BOOL := FALSE;
    StartCommandStack : BOOL := FALSE;
END_VAR

IF (SFCInit OR SFCReset) THEN
    CraneDown := FALSE;
    CraneOnConveyor := FALSE;
    CraneOnStack := FALSE;
    CraneSucked := FALSE;
    CraneUp := FALSE;
    StackGreenLamp := FALSE;
    StackSlider := FALSE;
    SFCInit := FALSE;
    SFCReset := FALSE;
    SliderMovedOut := FALSE;
    SliderNotMovedOut := FALSE;
    StartButtonStack := FALSE;
    StartCommandStack := FALSE;
    StartVar := FALSE;
    WorkpieceReady := FALSE;
    StackState := StackStates#StackSFCInit;
    interconnectStackStartCommand := FALSE;
END_IF;

IF NOT (SFCInit OR SFCPause) THEN
    CASE StackState OF
        StackStates#StackSFCInit:
            IF TRUE THEN
                StackState := StackStates#StartStack;
            END_IF;

        StackStates#StartStack:
            StackSlider := FALSE;
            StackGreenLamp := FALSE;
            StartVar := FALSE;
            StartCommandStack := FALSE;
            IF (StartButtonStack = TRUE) THEN
                interconnectStackStartCommand := TRUE;
            END_IF;
            IF interconnectStackStartCommand THEN
                StackState := StackStates#GreenLamp;
            END_IF;

        StackStates#GreenLamp:
            StackGreenLamp := TRUE;
            interconnectStackStartCommand := FALSE;
            IF TRUE THEN
                StackState := StackStates#StackInit;
            END_IF;

        StackStates#StackInit:
            StackSlider := TRUE;
            IF TRUE THEN
                StackState := StackStates#StackInit2;
            END_IF;

        StackStates#StackInit2:
            StackSlider := FALSE;
            IF TRUE THEN
                StackState := StackStates#Interstep;
            END_IF;

        StackStates#Interstep:
            StartCommandStack := TRUE;
            IF StartVar THEN
                StackState := StackStates#convey;
            END_IF;

        StackStates#convey:
            IF SliderNotMovedOut THEN
                StackSlider := TRUE;
            END_IF;
            IF CraneOnStack THEN
                StackState := StackStates#Step0;
            END_IF;

        StackStates#Step0:
            IF CraneDown THEN
                StackState := StackStates#SliderMoveBack;
            END_IF;

        StackStates#SliderMoveBack:
            IF ((SliderMovedOut = TRUE) AND (SliderNotMovedOut = FALSE)) THEN
                StackSlider := FALSE;
            END_IF;
            IF CraneUp THEN
                StackState := StackStates#Step1;
            END_IF;

        StackStates#Step1:
            IF CraneOnConveyor THEN
                StackState := StackStates#Interstep;
            END_IF;
    END_CASE;
END_IF;
END_FUNCTION_BLOCK

PROGRAM Main
VAR_INPUT
    SensorCraneDown : BOOL := FALSE;
    SensorCraneOnConveyor : BOOL := FALSE;
    SensorCraneOnStack : BOOL := FALSE;
    SensorCranePosition : BOOL := FALSE;
    SensorCraneSucked : BOOL := FALSE;
    SensorCraneUp : BOOL := FALSE;
    SensorStackEmergencyStop : BOOL := FALSE;
    SensorStackSwitchManuellAutomatic : BOOL := FALSE;
    SensorSliderMovedOut : BOOL := FALSE;
    SensorSliderNotMovedOut : BOOL := FALSE;
    SensorStartButtonStack : BOOL := FALSE;
    SensorWorkpieceReady : BOOL := FALSE;
END_VAR
VAR
    Crane : Crane;
    Stack : Stack;
END_VAR
VAR_OUTPUT
    ActuatorCraneLower : BOOL := FALSE;
    ActuatorCraneTurnClockwise : BOOL := FALSE;
    ActuatorCraneTurnCounterClockwise : BOOL := FALSE;
    ActuatorStackGreenLamp : BOOL := FALSE;
    ActuatorStackSlider : BOOL := FALSE;
    ActuatorStackVacuumOff : BOOL := FALSE;
    ActuatorStackVacuumOn : BOOL := FALSE;
    ActuatorStackWhiteLamp : BOOL := FALSE;
END_VAR
Stack.SliderNotMovedOut := SensorSliderNotMovedOut;
Stack.SliderMovedOut := SensorSliderMovedOut;
Stack.CraneOnStack := SensorCraneOnStack;
Stack.CraneDown := SensorCraneDown;
Stack.CraneUp := SensorCraneUp;
Stack.CraneOnConveyor := SensorCraneOnConveyor;
Stack.WorkpieceReady := SensorWorkpieceReady;
Stack.StartButtonStack := SensorStartButtonStack;
ActuatorStackSlider := Stack.StackSlider;
ActuatorStackGreenLamp := Stack.StackGreenLamp;
Crane.WorkpieceReady := SensorWorkpieceReady;
Crane.CraneUp := SensorCraneUp;
Crane.CraneOnConveyor := SensorCraneOnConveyor;
Crane.CraneDown := SensorCraneDown;
Crane.CraneSucked := SensorCraneSucked;
Crane.CraneOnStack := SensorCraneOnStack;
Crane.SliderMovedOut := SensorSliderMovedOut;
Crane.StartButtonStack := SensorStartButtonStack;
ActuatorCraneTurnCounterClockwise := Crane.CraneTurnCounterClockwise;
ActuatorCraneTurnClockwise := Crane.CraneTurnClockwise;
ActuatorCraneLower := Crane.CraneLower;
ActuatorStackVacuumOff := Crane.StackVacuumOff;
ActuatorStackVacuumOn := Crane.StackVacuumOn;
IF SensorStackEmergencyStop THEN
    Stack();
    Crane();
    IF ActuatorStackGreenLamp THEN
        IF (Crane.StartCommandCrane AND Stack.StartCommandStack) THEN
            Crane.StartVar := TRUE;
            Stack.StartVar := TRUE;
        END_IF;
    END_IF;
    Crane.SFCReset := FALSE;
    Stack.SFCReset := FALSE;
ELSIF NOT SensorStackEmergencyStop THEN
    ActuatorStackSlider := FALSE;
    ActuatorCraneLower := FALSE;
    ActuatorStackVacuumOn := FALSE;
    ActuatorStackVacuumOff := TRUE;
    ActuatorStackGreenLamp := FALSE;
    ActuatorCraneTurnCounterClockwise := FALSE;
    ActuatorCraneTurnClockwise := FALSE;
    Crane.SFCReset := TRUE;
    Stack.SFCReset := TRUE;
    Crane.StartVar := FALSE;
    Stack.StartVar := FALSE;
END_IF;
END_PROGRAM

FUNCTION_BLOCK TON
VAR_INPUT
    IN : BOOL;
    PT : TIME;
END_VAR
VAR
    running : BOOL;
END_VAR
VAR_TEMP
    timeout : BOOL;
END_VAR
VAR_OUTPUT
    Q : BOOL;
    ET : TIME;
END_VAR
timeout := NONDETERMINISTIC_BOOL();
IF NOT IN THEN
    Q := FALSE;
    running := FALSE;
ELSIF NOT running AND NOT Q THEN
    running := TRUE;
ELSIF running AND NOT Q THEN
    Q := timeout;
    running := NOT Q;
END_IF;
ET := NONDETERMINISTIC_TIME();
END_FUNCTION_BLOCK

(* ---- Scenario2_Final.st ---- *)
TYPE
    CraneStates : (CraneSFCInit, StartCrane, CraneInit, CraneInit2, Interstep, Interstep2, TimeDelay, TurnRight,
                   InterstepCheckWorkpiece, StackStop, Step0, CraneLiftStack, CraneTurnLeftNOTMetallic,
                   CraneOnConveyorState, CraneLiftStackMetallic, CraneTurnLeftMetallic, CraneOnConveyorMetallic,
                   release, CraneLiftConveyor, CraneStop);
    StackStates : (StackSFCInit, StartStack, GreenLamp, StackInit, StackInit2, Interstep, convey, Step0, SliderMoveBack,
                   Step1);
END_TYPE

FUNCTION_BLOCK Crane
VAR_INPUT
    CraneDown : BOOL := FALSE;
    CraneOnConveyor : BOOL := FALSE;
    CraneOnStack : BOOL := FALSE;
    CraneSucked : BOOL := FALSE;
    CraneUp : BOOL := FALSE;
    StackCapacitiveSensor : BOOL := FALSE;
    SFCReset : BOOL := FALSE;
    SliderMovedOut : BOOL := FALSE;
    SliderNotMovedOut : BOOL := FALSE;
    StartButtonStack : BOOL := FALSE;
    StartVar : BOOL := FALSE;
    WorkpieceReady : BOOL := FALSE;
END_VAR
VAR
    SFCInit : BOOL := FALSE;
    SFCPause : BOOL := FALSE;
    CraneState : CraneStates := CraneStates#CraneSFCInit;
    Timer : TON;
    TimerDuration : TIME := TIME#50.0ms;
    Timerinterconnect : BOOL := FALSE;
    interconnectCraneStartCommand : BOOL := FALSE;
END_VAR
VAR_OUTPUT
    CraneLower : BOOL := FALSE;
    CraneTurnClockwise : BOOL := FALSE;
    CraneTurnCounterClockwise : BOOL := FALSE;
    StackVacuumOff : BOOL := FALSE;
    StackVacuumOn : BOOL := FALSE;
    StartCommandCrane : BOOL := FALSE;
END_VAR

IF (SFCInit OR SFCReset) THEN
    CraneDown := FALSE;
    CraneLower := FALSE;
    CraneOnConveyor := FALSE;
    CraneOnStack := FALSE;
    CraneSucked := FALSE;
    CraneTurnClockwise := FALSE;
    CraneTurnCounterClockwise := FALSE;
    CraneUp := FALSE;
    StackCapacitiveSensor := FALSE;
    StackVacuumOff := FALSE;
    StackVacuumOn := FALSE;
    SFCInit := FALSE;
    SFCReset := FALSE;
    SliderMovedOut := FALSE;
    SliderNotMovedOut := FALSE;
    StartButtonStack := FALSE;
    StartCommandCrane := FALSE;
    StartVar := FALSE;
    Timer.ET := INT#0;
    Timer.IN := FALSE;
    Timer.PT := INT#0;
    Timer.Q := FALSE;
    TimerDuration := TIME#50ms;
    Timerinterconnect := FALSE;
    WorkpieceReady := FALSE;
    CraneState := CraneStates#CraneSFCInit;
    interconnectCraneStartCommand := FALSE;
END_IF;

IF NOT (SFCInit OR SFCPause) THEN
    CASE CraneState OF
        CraneStates#CraneSFCInit:
            IF TRUE THEN
                CraneState := CraneStates#StartCrane;
            END_IF;

        CraneStates#StartCrane:
            CraneLower := FALSE;
            StackVacuumOff := TRUE;
            StackVacuumOn := FALSE;
            CraneTurnCounterClockwise := FALSE;
            CraneTurnClockwise := FALSE;
            StartVar := FALSE;
            StartCommandCrane := FALSE;
            IF (StartButtonStack = TRUE) THEN
                interconnectCraneStartCommand := TRUE;
            END_IF;
            IF interconnectCraneStartCommand THEN
                CraneState := CraneStates#CraneInit;
            END_IF;

        CraneStates#CraneInit:
            CraneLower := TRUE;
            interconnectCraneStartCommand := FALSE;
            IF CraneDown THEN
                CraneState := CraneStates#CraneInit2;
            END_IF;

        CraneStates#CraneInit2:
            CraneLower := FALSE;
            IF CraneUp THEN
                CraneState := CraneStates#Interstep;
            END_IF;

        CraneStates#Interstep:
            StartCommandCrane := TRUE;
            IF StartVar THEN
                CraneState := CraneStates#Interstep2;
            END_IF;

        CraneStates#Interstep2:
            IF SliderMovedOut THEN
                CraneState := CraneStates#TimeDelay;
            END_IF;

        CraneStates#TimeDelay:
            Timer(IN := TRUE, PT := TimerDuration);
            Timerinterconnect := Timer.Q;
            IF Timerinterconnect THEN
                CraneState := CraneStates#TurnRight;
            END_IF;

        CraneStates#TurnRight:
            CraneTurnClockwise := TRUE;
            CraneTurnCounterClockwise := FALSE;
            IF CraneOnStack THEN
                CraneState := CraneStates#InterstepCheckWorkpiece;
            END_IF;

        CraneStates#InterstepCheckWorkpiece:
            IF WorkpieceReady THEN
                CraneState := CraneStates#StackStop;
            ELSIF NOT WorkpieceReady THEN
                CraneState := CraneStates#CraneStop;
            END_IF;

        CraneStates#StackStop:
            CraneTurnClockwise := FALSE;
            CraneTurnCounterClockwise := FALSE;
            StackVacuumOn := TRUE;
            StackVacuumOff := FALSE;
            CraneLower := TRUE;
            IF CraneSucked THEN
                CraneState := CraneStates#Step0;
            END_IF;

        CraneStates#Step0:
            IF NOT StackCapacitiveSensor THEN
                CraneState := CraneStates#CraneLiftStack;
            ELSIF StackCapacitiveSensor THEN
                CraneState := CraneStates#CraneLiftStackMetallic;
            END_IF;

        CraneStates#CraneLiftStack:
            CraneLower := FALSE;
            IF CraneUp THEN
                CraneState := CraneStates#CraneTurnLeftNOTMetallic;
            END_IF;

        CraneStates#CraneTurnLeftNOTMetallic:
            CraneTurnCounterClockwise := TRUE;
            CraneTurnClockwise := FALSE;
            IF CraneOnConveyor THEN
                CraneState := CraneStates#CraneOnConveyorState;
            END_IF;

        CraneStates#CraneOnConveyorState:
            CraneTurnCounterClockwise := FALSE;
            CraneTurnClockwise := FALSE;
            CraneLower := TRUE;
            IF CraneDown THEN
                CraneState := CraneStates#release;
            END_IF;

        CraneStates#CraneLiftStackMetallic:
            CraneLower := FALSE;
            IF CraneUp THEN
                CraneState := CraneStates#CraneTurnLeftMetallic;
            END_IF;

        CraneStates#CraneTurnLeftMetallic:
            CraneTurnCounterClockwise := TRUE;
            CraneTurnClockwise := FALSE;
            IF CraneOnConveyor THEN
                CraneState := CraneStates#CraneOnConveyorMetallic;
            END_IF;

        CraneStates#CraneOnConveyorMetallic:
            CraneTurnCounterClockwise := FALSE;
            CraneTurnClockwise := FALSE;
            CraneLower := TRUE;
            IF CraneDown THEN
                CraneState := CraneStates#release;
            END_IF;

        CraneStates#release:
            StackVacuumOff := TRUE;
            StackVacuumOn := FALSE;
            IF TRUE THEN
                CraneState := CraneStates#CraneLiftConveyor;
            END_IF;

        CraneStates#CraneLiftConveyor:
            CraneLower := FALSE;
            IF TRUE THEN
                CraneState := CraneStates#Interstep;
            END_IF;

        CraneStates#CraneStop:
            IF TRUE THEN
                CraneState := CraneStates#StartCrane;
            END_IF;
    END_CASE;
END_IF;
END_FUNCTION_BLOCK

FUNCTION_BLOCK Stack
VAR_INPUT
    CraneDown : BOOL := FALSE;
    CraneOnConveyor : BOOL := FALSE;
    CraneOnStack : BOOL := FALSE;
    CraneSucked : BOOL := FALSE;
    CraneUp : BOOL := FALSE;
    SFCReset : BOOL := FALSE;
    SliderMovedOut : BOOL := FALSE;
    SliderNotMovedOut : BOOL := FALSE;
    StartButtonStack : BOOL := FALSE;
    StartVar : BOOL := FALSE;
    WorkpieceReady : BOOL := FALSE;
END_VAR
VAR
    SFCInit : BOOL := FALSE;
    SFCPause : BOOL := FALSE;
    StackState : StackStates := StackStates#StackSFCInit;
    interconnectStackStartCommand : BOOL := FALSE;
END_VAR
VAR_OUTPUT
    CraneLower : BOOL := FALSE;
    CraneTurnClockwise : BOOL := FALSE;
    CraneTurnCounterClockwise : BOOL := FALSE;
    StackGreenLamp : BOOL := FALSE;
    StackSlider : BOOL := FALSE;
    StackVacuumOff : BOOL := FALSE;
    StackVacuumOn : BOOL := FALSE;
    StackWhiteLamp : BOOL := FALSE;
    StartCommandStack : BOOL := FALSE;
END_VAR

IF (SFCInit OR SFCReset) THEN
    CraneDown := FALSE;
    CraneLower := FALSE;
    CraneOnConveyor := FALSE;
    CraneOnStack := FALSE;
    CraneSucked := FALSE;
    CraneTurnClockwise := FALSE;
    CraneTurnCounterClockwise := FALSE;
    CraneUp := FALSE;
    StackGreenLamp := FALSE;
    StackSlider := FALSE;
    StackVacuumOff := FALSE;
    StackVacuumOn := FALSE;
    StackWhiteLamp := FALSE;
    SFCInit := FALSE;
    SFCReset := FALSE;
    SliderMovedOut := FALSE;
    SliderNotMovedOut := FALSE;
    StartButtonStack := FALSE;
    StartCommandStack := FALSE;
    StartVar := FALSE;
    WorkpieceReady := FALSE;
    StackState := StackStates#StackSFCInit;
    interconnectStackStartCommand := FALSE;
END_IF;

IF NOT (SFCInit OR SFCPause) THEN
    CASE StackState OF
        StackStates#StackSFCInit:
            IF TRUE THEN
                StackState := StackStates#StartStack;
            END_IF;

        StackStates#StartStack:
            StackSlider := FALSE;
            StackGreenLamp := FALSE;
            StartVar := FALSE;
            StartCommandStack := FALSE;
            IF (StartButtonStack = TRUE) THEN
                interconnectStackStartCommand := TRUE;
            END_IF;
            IF interconnectStackStartCommand THEN
                StackState := StackStates#GreenLamp;
            END_IF;

        StackStates#GreenLamp:
            StackGreenLamp := TRUE;
            interconnectStackStartCommand := FALSE;
            IF TRUE THEN
                StackState := StackStates#StackInit;
            END_IF;

        StackStates#StackInit:
            StackSlider := TRUE;
            IF TRUE THEN
                StackState := StackStates#StackInit2;
            END_IF;

        StackStates#StackInit2:
            StackSlider := FALSE;
            IF TRUE THEN
                StackState := StackStates#Interstep;
            END_IF;

        StackStates#Interstep:
            StartCommandStack := TRUE;
            IF StartVar THEN
                StackState := StackStates#convey;
            END_IF;

        StackStates#convey:
            IF SliderNotMovedOut THEN
                StackSlider := TRUE;
            END_IF;
            IF CraneOnStack THEN
                StackState := StackStates#Step0;
            END_IF;

        StackStates#Step0:
            IF CraneDown THEN
                StackState := StackStates#SliderMoveBack;
            END_IF;

        StackStates#SliderMoveBack:
            IF ((SliderMovedOut = TRUE) AND (SliderNotMovedOut = FALSE)) THEN
                StackSlider := FALSE;
            END_IF;
            IF CraneUp THEN
                StackState := StackStates#Step1;
            END_IF;

        StackStates#Step1:
            IF CraneOnConveyor THEN
                StackState := StackStates#Interstep;
            END_IF;
    END_CASE;
END_IF;
END_FUNCTION_BLOCK

PROGRAM Main
VAR_INPUT
    SensorCraneDown : BOOL := FALSE;
    SensorCraneOnConveyor : BOOL := FALSE;
    SensorCraneOnStack : BOOL := FALSE;
    SensorCranePosition : BOOL := FALSE;
    SensorCranePositionStamp : BOOL := FALSE;
    SensorCraneSucked : BOOL := FALSE;
    SensorCraneUp : BOOL := FALSE;
    SensorStackCapacitiveSensor : BOOL := FALSE;
    SensorStackEmergencyStop : BOOL := FALSE;
    SensorStackOpticalSensor : BOOL := FALSE;
    SensorStackSwitchManuellAutomatic : BOOL := FALSE;
    SensorSliderMovedOut : BOOL := FALSE;
    SensorSliderNotMovedOut : BOOL := FALSE;
    SensorStartButtonStack : BOOL := FALSE;
    SensorWorkpieceReady : BOOL := FALSE;
END_VAR
VAR
    Crane : Crane;
    Stack : Stack;
END_VAR
VAR_OUTPUT
    ActuatorCraneLower : BOOL := FALSE;
    ActuatorCraneTurnClockwise : BOOL := FALSE;
    ActuatorCraneTurnCounterClockwise : BOOL := FALSE;
    ActuatorStackGreenLamp : BOOL := FALSE;
    ActuatorStackSlider : BOOL := FALSE;
    ActuatorStackVacuumOff : BOOL := FALSE;
    ActuatorStackVacuumOn : BOOL := FALSE;
    ActuatorStackWhiteLamp : BOOL := FALSE;
END_VAR
Stack.SliderNotMovedOut := SensorSliderNotMovedOut;
Stack.SliderMovedOut := SensorSliderMovedOut;
Stack.CraneOnStack := SensorCraneOnStack;
Stack.CraneDown := SensorCraneDown;
Stack.CraneUp := SensorCraneUp;
Stack.CraneOnConveyor := SensorCraneOnConveyor;
Stack.WorkpieceReady := SensorWorkpieceReady;
Stack.StartButtonStack := SensorStartButtonStack;
ActuatorStackSlider := Stack.StackSlider;
ActuatorStackGreenLamp := Stack.StackGreenLamp;
Crane.WorkpieceReady := SensorWorkpieceReady;
Crane.CraneUp := SensorCraneUp;
Crane.CraneOnConveyor := SensorCraneOnConveyor;
Crane.CraneDown := SensorCraneDown;
Crane.CraneSucked := SensorCraneSucked;
Crane.CraneOnStack := SensorCraneOnStack;
Crane.StackCapacitiveSensor := SensorStackCapacitiveSensor;
Crane.SliderMovedOut := SensorSliderMovedOut;
Crane.StartButtonStack := SensorStartButtonStack;
ActuatorCraneTurnCounterClockwise := Crane.CraneTurnCounterClockwise;
ActuatorCraneTurnClockwise := Crane.CraneTurnClockwise;
ActuatorCraneLower := Crane.CraneLower;
ActuatorStackVacuumOff := Crane.StackVacuumOff;
ActuatorStackVacuumOn := Crane.StackVacuumOn;
IF SensorStackEmergencyStop THEN
    Stack();
    Crane();
    IF ActuatorStackGreenLamp THEN
        IF (Crane.StartCommandCrane AND Stack.StartCommandStack) THEN
            Crane.StartVar := TRUE;
            Stack.StartVar := TRUE;
        END_IF;
    END_IF;
    Crane.SFCReset := FALSE;
    Stack.SFCReset := FALSE;
ELSIF NOT SensorStackEmergencyStop THEN
    ActuatorStackSlider := FALSE;
    ActuatorCraneLower := FALSE;
    ActuatorStackVacuumOn := FALSE;
    ActuatorStackVacuumOff := TRUE;
    ActuatorStackGreenLamp := FALSE;
    ActuatorCraneTurnCounterClockwise := FALSE;
    ActuatorCraneTurnClockwise := FALSE;
    Crane.SFCReset := TRUE;
    Stack.SFCReset := TRUE;
    Crane.StartVar := FALSE;
    Stack.StartVar := FALSE;
END_IF;
END_PROGRAM

FUNCTION_BLOCK TON
VAR_INPUT
    IN : BOOL;
    PT : TIME;
END_VAR
VAR
    running : BOOL;
END_VAR
VAR_TEMP
    timeout : BOOL;
END_VAR
VAR_OUTPUT
    Q : BOOL;
    ET : TIME;
END_VAR
timeout := NONDETERMINISTIC_BOOL();
IF NOT IN THEN
    Q := FALSE;
    running := FALSE;
ELSIF NOT running AND NOT Q THEN
    running := TRUE;
ELSIF running AND NOT Q THEN
    Q := timeout;
    running := NOT Q;
END_IF;
ET := NONDETERMINISTIC_TIME();
END_FUNCTION_BLOCK

(* ---- Scenario3_Final.st ---- *)
TYPE
    CraneStates : (CraneSFCInit, StartCrane, CraneInit, CraneInit2, Interstep, Interstep2, TimeDelay, TurnRight,
                   InterstepCheckWorkpiece, StackStop, Step0, CraneLiftStack, CraneTurnLeftNOTMetallic,
                   CraneOnConveyorState, CraneLiftStackMetallic, CraneTurnLeftMetallic, CraneOnStampMetallic,
                   releaseWorkpiece, CraneGoUp, pause, Resetinterconnect, LowerCrane, SuckAtStamp, CraneLiftAtStamp,
                   CraneTurnLeftFromStamp, CraneOnConveyorMetallic, release, CraneLiftConveyor, WaitAtStamp, Step2);
    StackStates : (StackSFCInit, StartStack, GreenLamp, StackInit, StackInit2, Interstep, convey, Step0, SliderMoveBack,
                   Step1);
    StampStates : (StampSFCInit, StartStamp, GreenLamp, StampInit1, StampInit2, StampInit3, StampInit4, Interstep,
                   Interstep2, Step0, StampSliderBack, StampProcess, Step1, StampSliderForward, Step2);
END_TYPE

FUNCTION_BLOCK Crane
VAR_INPUT
    CraneDown : BOOL := FALSE;
    CraneOnConveyor : BOOL := FALSE;
    CraneOnStack : BOOL := FALSE;
    CranePositionStamp : BOOL := FALSE;
    CraneSucked : BOOL := FALSE;
    CraneUp : BOOL := FALSE;
    StackCapacitiveSensor : BOOL := FALSE;
    SFCReset : BOOL := FALSE;
    SliderMovedOut : BOOL := FALSE;
    SliderNotMovedOut : BOOL := FALSE;
    StampLowered : BOOL := FALSE;
    StampSliderFilled : BOOL := FALSE;
    StartButtonStack : BOOL := FALSE;
    StartVar : BOOL := FALSE;
    WorkpieceReady : BOOL := FALSE;
END_VAR
VAR
    Duration1 : TIME := TIME#1500.0ms;
    SFCInit : BOOL := FALSE;
    SFCPause : BOOL := FALSE;
    CraneState : CraneStates := CraneStates#CraneSFCInit;
    Timer : TON;
    TimerDuration : TIME := TIME#50.0ms;
    Timerinterconnect : BOOL := FALSE;
    Timer1 : TON;
    interconnect : BOOL := FALSE;
    interconnectCraneStartCommand : BOOL := FALSE;
END_VAR
VAR_OUTPUT
    CraneLower : BOOL := FALSE;
    CraneTurnClockwise : BOOL := FALSE;
    CraneTurnCounterClockwise : BOOL := FALSE;
    StackVacuumOff : BOOL := FALSE;
    StackVacuumOn : BOOL := FALSE;
    StartCommandCrane : BOOL := FALSE;
END_VAR

IF (SFCInit OR SFCReset) THEN
    CraneDown := FALSE;
    CraneLower := FALSE;
    CraneOnConveyor := FALSE;
    CraneOnStack := FALSE;
    CranePositionStamp := FALSE;
    CraneSucked := FALSE;
    CraneTurnClockwise := FALSE;
    CraneTurnCounterClockwise := FALSE;
    CraneUp := FALSE;
    Duration1 := TIME#1500ms;
    StackCapacitiveSensor := FALSE;
    StackVacuumOff := FALSE;
    StackVacuumOn := FALSE;
    SFCInit := FALSE;
    SFCReset := FALSE;
    SliderMovedOut := FALSE;
    SliderNotMovedOut := FALSE;
    StampLowered := FALSE;
    StampSliderFilled := FALSE;
    StartButtonStack := FALSE;
    StartCommandCrane := FALSE;
    StartVar := FALSE;
    Timer.ET := INT#0;
    Timer.IN := FALSE;
    Timer.PT := INT#0;
    Timer.Q := FALSE;
    TimerDuration := TIME#50ms;
    Timerinterconnect := FALSE;
    Timer1.ET := INT#0;
    Timer1.IN := FALSE;
    Timer1.PT := INT#0;
    Timer1.Q := FALSE;
    WorkpieceReady := FALSE;
    CraneState := CraneStates#CraneSFCInit;
    interconnect := FALSE;
    interconnectCraneStartCommand := FALSE;
END_IF;

IF NOT (SFCInit OR SFCPause) THEN
    CASE CraneState OF
        CraneStates#CraneSFCInit:
            IF TRUE THEN
                CraneState := CraneStates#StartCrane;
            END_IF;

        CraneStates#StartCrane:
            CraneLower := FALSE;
            StackVacuumOff := TRUE;
            StackVacuumOn := FALSE;
            CraneTurnCounterClockwise := FALSE;
            CraneTurnClockwise := FALSE;
            StartVar := FALSE;
            StartCommandCrane := FALSE;
            IF (StartButtonStack = TRUE) THEN
                interconnectCraneStartCommand := TRUE;
            END_IF;
            IF interconnectCraneStartCommand THEN
                CraneState := CraneStates#CraneInit;
            END_IF;

        CraneStates#CraneInit:
            CraneLower := TRUE;
            interconnectCraneStartCommand := FALSE;
            IF CraneDown THEN
                CraneState := CraneStates#CraneInit2;
            END_IF;

        CraneStates#CraneInit2:
            CraneLower := FALSE;
            IF CraneUp THEN
                CraneState := CraneStates#Interstep;
            END_IF;

        CraneStates#Interstep:
            StartCommandCrane := TRUE;
            IF StartVar THEN
                CraneState := CraneStates#Interstep2;
            END_IF;

        CraneStates#Interstep2:
            IF SliderMovedOut THEN
                CraneState := CraneStates#TimeDelay;
            END_IF;

        CraneStates#TimeDelay:
            Timer(IN := TRUE, PT := TimerDuration);
            Timerinterconnect := Timer.Q;
            IF Timerinterconnect THEN
                CraneState := CraneStates#TurnRight;
            END_IF;

        CraneStates#TurnRight:
            CraneTurnClockwise := TRUE;
            CraneTurnCounterClockwise := FALSE;
            IF CraneOnStack THEN
                CraneState := CraneStates#InterstepCheckWorkpiece;
            END_IF;

        CraneStates#InterstepCheckWorkpiece:
            IF WorkpieceReady THEN
                CraneState := CraneStates#StackStop;
            ELSIF (NOT WorkpieceReady AND StampSliderFilled) THEN
                CraneState := CraneStates#WaitAtStamp;
            ELSIF (NOT WorkpieceReady AND NOT StampSliderFilled) THEN
                CraneState := CraneStates#Step2;
            END_IF;

        CraneStates#StackStop:
            CraneTurnClockwise := FALSE;
            CraneTurnCounterClockwise := FALSE;
            StackVacuumOn := TRUE;
            StackVacuumOff := FALSE;
            CraneLower := TRUE;
            IF CraneSucked THEN
                CraneState := CraneStates#Step0;
            END_IF;

        CraneStates#Step0:
            IF NOT StackCapacitiveSensor THEN
                CraneState := CraneStates#CraneLiftStack;
            ELSIF StackCapacitiveSensor THEN
                CraneState := CraneStates#CraneLiftStackMetallic;
            END_IF;

        CraneStates#CraneLiftStack:
            CraneLower := FALSE;
            IF CraneUp THEN
                CraneState := CraneStates#CraneTurnLeftNOTMetallic;
            END_IF;

        CraneStates#CraneTurnLeftNOTMetallic:
            CraneTurnCounterClockwise := TRUE;
            CraneTurnClockwise := FALSE;
            IF CraneOnConveyor THEN
                CraneState := CraneStates#CraneOnConveyorState;
            END_IF;

        CraneStates#CraneOnConveyorState:
            CraneTurnCounterClockwise := FALSE;
            CraneTurnClockwise := FALSE;
            CraneLower := TRUE;
            IF CraneDown THEN
                CraneState := CraneStates#release;
            END_IF;

        CraneStates#CraneLiftStackMetallic:
            CraneLower := FALSE;
            IF CraneUp THEN
                CraneState := CraneStates#CraneTurnLeftMetallic;
            END_IF;

        CraneStates#CraneTurnLeftMetallic:
            CraneTurnCounterClockwise := TRUE;
            CraneTurnClockwise := FALSE;
            IF CranePositionStamp THEN
                CraneState := CraneStates#CraneOnStampMetallic;
            END_IF;

        CraneStates#CraneOnStampMetallic:
            CraneTurnCounterClockwise := FALSE;
            CraneTurnClockwise := FALSE;
            CraneLower := TRUE;
            IF CraneDown THEN
                CraneState := CraneStates#releaseWorkpiece;
            END_IF;

        CraneStates#releaseWorkpiece:
            StackVacuumOff := TRUE;
            StackVacuumOn := FALSE;
            IF TRUE THEN
                CraneState := CraneStates#CraneGoUp;
            END_IF;

        CraneStates#CraneGoUp:
            CraneLower := FALSE;
            IF CraneUp THEN
                CraneState := CraneStates#pause;
            END_IF;

        CraneStates#pause:
            Timer1(IN := CraneUp, PT := Duration1);
            interconnect := Timer1.Q;
            IF interconnect THEN
                CraneState := CraneStates#Resetinterconnect;
            END_IF;

        CraneStates#Resetinterconnect:
            interconnect := FALSE;
            Timer1(IN := FALSE, PT := TIME#1ms);
            IF SliderMovedOut THEN
                CraneState := CraneStates#LowerCrane;
            END_IF;

        CraneStates#LowerCrane:
            CraneLower := TRUE;
            IF CraneDown THEN
                CraneState := CraneStates#SuckAtStamp;
            END_IF;

        CraneStates#SuckAtStamp:
            StackVacuumOn := TRUE;
            StackVacuumOff := FALSE;
            IF CraneSucked THEN
                CraneState := CraneStates#CraneLiftAtStamp;
            END_IF;

        CraneStates#CraneLiftAtStamp:
            CraneLower := FALSE;
            IF CraneUp THEN
                CraneState := CraneStates#CraneTurnLeftFromStamp;
            END_IF;

        CraneStates#CraneTurnLeftFromStamp:
            CraneTurnClockwise := TRUE;
            CraneTurnCounterClockwise := FALSE;
            IF CraneOnConveyor THEN
                CraneState := CraneStates#CraneOnConveyorMetallic;
            END_IF;

        CraneStates#CraneOnConveyorMetallic:
            CraneTurnCounterClockwise := FALSE;
            CraneTurnClockwise := FALSE;
            CraneLower := TRUE;
            IF CraneDown THEN
                CraneState := CraneStates#release;
            END_IF;

        CraneStates#release:
            StackVacuumOff := TRUE;
            StackVacuumOn := FALSE;
            IF TRUE THEN
                CraneState := CraneStates#CraneLiftConveyor;
            END_IF;

        CraneStates#CraneLiftConveyor:
            CraneLower := FALSE;
            IF TRUE THEN
                CraneState := CraneStates#Interstep;
            END_IF;

        CraneStates#WaitAtStamp:
            IF TRUE THEN
                CraneState := CraneStates#pause;
            END_IF;

        CraneStates#Step2:
            IF TRUE THEN
                CraneState := CraneStates#StartCrane;
            END_IF;
    END_CASE;
END_IF;
END_FUNCTION_BLOCK

FUNCTION_BLOCK Stack
VAR_INPUT
    CraneDown : BOOL := FALSE;
    CraneOnConveyor : BOOL := FALSE;
    CraneOnStack : BOOL := FALSE;
    CraneSucked : BOOL := FALSE;
    CraneUp : BOOL := FALSE;
    SFCReset : BOOL := FALSE;
    SliderMovedOut : BOOL := FALSE;
    SliderNotMovedOut : BOOL := FALSE;
    StartButtonStack : BOOL := FALSE;
    StartVar : BOOL := FALSE;
    WorkpieceReady : BOOL := FALSE;
END_VAR
VAR
    SFCInit : BOOL := FALSE;
    SFCPause : BOOL := FALSE;
    StackState : StackStates := StackStates#StackSFCInit;
    interconnectStackStartCommand : BOOL := FALSE;
END_VAR
VAR_OUTPUT
    CraneLower : BOOL := FALSE;
    CraneTurnClockwise : BOOL := FALSE;
    CraneTurnCounterClockwise : BOOL := FALSE;
    StackGreenLamp : BOOL := FALSE;
    StackSlider : BOOL := FALSE;
    StackVacuumOff : BOOL := FALSE;
    StackVacuumOn : BOOL := FALSE;
    StackWhiteLamp : BOOL := FALSE;
    StartCommandStack : BOOL := FALSE;
END_VAR

IF (SFCInit OR SFCReset) THEN
    CraneDown := FALSE;
    CraneLower := FALSE;
    CraneOnConveyor := FALSE;
    CraneOnStack := FALSE;
    CraneSucked := FALSE;
    CraneTurnClockwise := FALSE;
    CraneTurnCounterClockwise := FALSE;
    CraneUp := FALSE;
    StackGreenLamp := FALSE;
    StackSlider := FALSE;
    StackVacuumOff := FALSE;
    StackVacuumOn := FALSE;
    StackWhiteLamp := FALSE;
    SFCInit := FALSE;
    SFCReset := FALSE;
    SliderMovedOut := FALSE;
    SliderNotMovedOut := FALSE;
    StartButtonStack := FALSE;
    StartCommandStack := FALSE;
    StartVar := FALSE;
    WorkpieceReady := FALSE;
    StackState := StackStates#StackSFCInit;
    interconnectStackStartCommand := FALSE;
END_IF;

IF NOT (SFCInit OR SFCPause) THEN
    CASE StackState OF
        StackStates#StackSFCInit:
            IF TRUE THEN
                StackState := StackStates#StartStack;
            END_IF;

        StackStates#StartStack:
            StackSlider := FALSE;
            StackGreenLamp := FALSE;
            StartVar := FALSE;
            StartCommandStack := FALSE;
            IF (StartButtonStack = TRUE) THEN
                interconnectStackStartCommand := TRUE;
            END_IF;
            IF interconnectStackStartCommand THEN
                StackState := StackStates#GreenLamp;
            END_IF;

        StackStates#GreenLamp:
            StackGreenLamp := TRUE;
            interconnectStackStartCommand := FALSE;
            IF TRUE THEN
                StackState := StackStates#StackInit;
            END_IF;

        StackStates#StackInit:
            StackSlider := TRUE;
            IF TRUE THEN
                StackState := StackStates#StackInit2;
            END_IF;

        StackStates#StackInit2:
            StackSlider := FALSE;
            IF TRUE THEN
                StackState := StackStates#Interstep;
            END_IF;

        StackStates#Interstep:
            StartCommandStack := TRUE;
            IF StartVar THEN
                StackState := StackStates#convey;
            END_IF;

        StackStates#convey:
            IF SliderNotMovedOut THEN
                StackSlider := TRUE;
            END_IF;
            IF CraneOnStack THEN
                StackState := StackStates#Step0;
            END_IF;

        StackStates#Step0:
            IF CraneDown THEN
                StackState := StackStates#SliderMoveBack;
            END_IF;

        StackStates#SliderMoveBack:
            IF ((SliderMovedOut = TRUE) AND (SliderNotMovedOut = FALSE)) THEN
                StackSlider := FALSE;
            END_IF;
            IF CraneUp THEN
                StackState := StackStates#Step1;
            END_IF;

        StackStates#Step1:
            IF CraneOnConveyor THEN
                StackState := StackStates#Interstep;
            END_IF;
    END_CASE;
END_IF;
END_FUNCTION_BLOCK

FUNCTION_BLOCK Stamp
VAR_INPUT
    CraneDown : BOOL := FALSE;
    CraneOnConveyor : BOOL := FALSE;
    CranePositionStamp : BOOL := FALSE;
    CraneSucked : BOOL := FALSE;
    CraneUp : BOOL := FALSE;
    SFCReset : BOOL := FALSE;
    StampLowered : BOOL := FALSE;
    StampSliderFilled : BOOL := FALSE;
    StampSliderSensorMovedIn : BOOL := FALSE;
    StampSliderSensorMovedOut : BOOL := FALSE;
    StampStartButton : BOOL := FALSE;
    StampUp : BOOL := FALSE;
    StartVar : BOOL := FALSE;
END_VAR
VAR
    Duration : TIME := TIME#500.0ms;
    SFCInit : BOOL := FALSE;
    SFCPause : BOOL := FALSE;
    StampState : StampStates := StampStates#StampSFCInit;
    Timer : TON;
    interconnect : BOOL := FALSE;
    interconnectStampStartCommand : BOOL := FALSE;
END_VAR
VAR_OUTPUT
    StampGreenLamp : BOOL := FALSE;
    StampPressure : BOOL := FALSE;
    StampPusher : BOOL := FALSE;
    StampSliderMovedIn : BOOL := FALSE;
    StampSliderMovedOut : BOOL := FALSE;
    StampWhiteLamp : BOOL := FALSE;
    StartCommandStamp : BOOL := FALSE;
END_VAR

IF (SFCInit OR SFCReset) THEN
    CraneDown := FALSE;
    CraneOnConveyor := FALSE;
    CranePositionStamp := FALSE;
    CraneSucked := FALSE;
    CraneUp := FALSE;
    Duration := TIME#500ms;
    SFCInit := FALSE;
    SFCReset := FALSE;
    StampGreenLamp := FALSE;
    StampLowered := FALSE;
    StampPressure := FALSE;
    StampPusher := FALSE;
    StampSliderFilled := FALSE;
    StampSliderMovedIn := FALSE;
    StampSliderMovedOut := FALSE;
    StampSliderSensorMovedIn := FALSE;
    StampSliderSensorMovedOut := FALSE;
    StampStartButton := FALSE;
    StampUp := FALSE;
    StampWhiteLamp := FALSE;
    StartCommandStamp := FALSE;
    StartVar := FALSE;
    Timer.ET := INT#0;
    Timer.IN := FALSE;
    Timer.PT := INT#0;
    Timer.Q := FALSE;
    StampState := StampStates#StampSFCInit;
    interconnect := FALSE;
    interconnectStampStartCommand := FALSE;
END_IF;

IF NOT (SFCInit OR SFCPause) THEN
    CASE StampState OF
        StampStates#StampSFCInit:
            IF TRUE THEN
                StampState := StampStates#StartStamp;
            END_IF;

        StampStates#StartStamp:
            StampSliderMovedOut := FALSE;
            StampSliderMovedIn := FALSE;
            StampPusher := FALSE;
            StampGreenLamp := FALSE;
            StampPressure := FALSE;
            StartCommandStamp := FALSE;
            IF (StampStartButton = TRUE) THEN
                interconnectStampStartCommand := TRUE;
            END_IF;
            IF interconnectStampStartCommand THEN
                StampState := StampStates#GreenLamp;
            END_IF;

        StampStates#GreenLamp:
            StampGreenLamp := TRUE;
            interconnectStampStartCommand := FALSE;
            IF TRUE THEN
                StampState := StampStates#StampInit1;
            END_IF;

        StampStates#StampInit1:
            StampSliderMovedIn := TRUE;
            StampSliderMovedOut := FALSE;
            IF StampSliderSensorMovedIn THEN
                StampState := StampStates#StampInit2;
            END_IF;

        StampStates#StampInit2:
            StampSliderMovedIn := FALSE;
            StampSliderMovedOut := TRUE;
            IF StampSliderSensorMovedOut THEN
                StampState := StampStates#StampInit3;
            END_IF;

        StampStates#StampInit3:
            StampPusher := TRUE;
            IF StampLowered THEN
                StampState := StampStates#StampInit4;
            END_IF;

        StampStates#StampInit4:
            StampPusher := FALSE;
            IF StampUp THEN
                StampState := StampStates#Interstep;
            END_IF;

        StampStates#Interstep:
            StartCommandStamp := TRUE;
            IF StartVar THEN
                StampState := StampStates#Interstep2;
            END_IF;

        StampStates#Interstep2:
            IF StampSliderFilled THEN
                StampState := StampStates#Step0;
            END_IF;

        StampStates#Step0:
            IF CraneUp THEN
                StampState := StampStates#StampSliderBack;
            END_IF;

        StampStates#StampSliderBack:
            StampSliderMovedIn := TRUE;
            StampSliderMovedOut := FALSE;
            IF StampSliderSensorMovedIn THEN
                StampState := StampStates#StampProcess;
            END_IF;

        StampStates#StampProcess:
            StampSliderMovedIn := FALSE;
            StampPusher := TRUE;
            IF StampLowered THEN
                StampState := StampStates#Step1;
            END_IF;

        StampStates#Step1:
            Timer(IN := StampLowered, PT := TIME#0ms);
            interconnect := Timer.Q;
            IF interconnect THEN
                StampState := StampStates#StampSliderForward;
            END_IF;

        StampStates#StampSliderForward:
            StampPusher := FALSE;
            StampSliderMovedOut := TRUE;
            IF ((StampLowered = FALSE) AND (StampUp = TRUE)) THEN
                interconnect := FALSE;
            END_IF;
            Timer(IN := FALSE, PT := TIME#1ms);
            IF StampSliderMovedOut THEN
                StampState := StampStates#Step2;
            END_IF;

        StampStates#Step2:
            IF CraneOnConveyor THEN
                StampState := StampStates#Interstep;
            END_IF;
    END_CASE;
END_IF;
END_FUNCTION_BLOCK

PROGRAM Main
VAR_INPUT
    SensorCraneDown : BOOL := FALSE;
    SensorCraneOnConveyor : BOOL := FALSE;
    SensorCraneOnStack : BOOL := FALSE;
    SensorCranePosition : BOOL := FALSE;
    SensorCranePositionStamp : BOOL := FALSE;
    SensorCraneSucked : BOOL := FALSE;
    SensorCraneUp : BOOL := FALSE;
    SensorStackCapacitiveSensor : BOOL := FALSE;
    SensorStackEmergencyStop : BOOL := FALSE;
    SensorStackOpticalSensor : BOOL := FALSE;
    SensorStackSwitchManuellAutomatic : BOOL := FALSE;
    SensorSliderMovedOut : BOOL := FALSE;
    SensorSliderNotMovedOut : BOOL := FALSE;
    SensorStampEmergencyStop : BOOL := FALSE;
    SensorStampLowered : BOOL := FALSE;
    SensorStampSliderFilled : BOOL := FALSE;
    SensorStampSliderSensorMovedIn : BOOL := FALSE;
    SensorStampSliderSensorMovedOut : BOOL := FALSE;
    SensorStampStartButton : BOOL := FALSE;
    SensorStampSwitchManuellAutomatic : BOOL := FALSE;
    SensorStampUp : BOOL := FALSE;
    SensorStartButtonStack : BOOL := FALSE;
    SensorWorkpieceReady : BOOL := FALSE;
END_VAR
VAR
    Crane : Crane;
    Stack : Stack;
    Stamp : Stamp;
END_VAR
VAR_OUTPUT
    ActuatorAnalogCranePressure : INT := 0;
    ActuatorCraneLower : BOOL := FALSE;
    ActuatorCraneTurnClockwise : BOOL := FALSE;
    ActuatorCraneTurnCounterClockwise : BOOL := FALSE;
    ActuatorStackGreenLamp : BOOL := FALSE;
    ActuatorStackSlider : BOOL := FALSE;
    ActuatorStackVacuumOff : BOOL := FALSE;
    ActuatorStackVacuumOn : BOOL := FALSE;
    ActuatorStackWhiteLamp : BOOL := FALSE;
    ActuatorSomeActuator : BOOL := FALSE;
    ActuatorStampGreenLamp : BOOL := FALSE;
    ActuatorStampPusher : BOOL := FALSE;
    ActuatorStampSliderMovedIn : BOOL := FALSE;
    ActuatorStampSliderMovedOut : BOOL := FALSE;
    ActuatorStampWhiteLamp : BOOL := FALSE;
END_VAR
Stack.SliderNotMovedOut := SensorSliderNotMovedOut;
Stack.SliderMovedOut := SensorSliderMovedOut;
Stack.CraneOnStack := SensorCraneOnStack;
Stack.CraneDown := SensorCraneDown;
Stack.CraneUp := SensorCraneUp;
Stack.CraneOnConveyor := SensorCraneOnConveyor;
Stack.WorkpieceReady := SensorWorkpieceReady;
Stack.StartButtonStack := SensorStartButtonStack;
ActuatorStackSlider := Stack.StackSlider;
ActuatorStackGreenLamp := Stack.StackGreenLamp;
Crane.CraneUp := SensorCraneUp;
Crane.CraneOnConveyor := SensorCraneOnConveyor;
Crane.CraneDown := SensorCraneDown;
Crane.CraneSucked := SensorCraneSucked;
Crane.CraneOnStack := SensorCraneOnStack;
Crane.StackCapacitiveSensor := SensorStackCapacitiveSensor;
Crane.CranePositionStamp := SensorCranePositionStamp;
Crane.SliderMovedOut := SensorSliderMovedOut;
Crane.WorkpieceReady := SensorWorkpieceReady;
Crane.StampSliderFilled := SensorStampSliderFilled;
Crane.SliderMovedOut := SensorSliderMovedOut;
Crane.StartButtonStack := SensorStartButtonStack;
ActuatorCraneTurnCounterClockwise := Crane.CraneTurnCounterClockwise;
ActuatorCraneTurnClockwise := Crane.CraneTurnClockwise;
ActuatorCraneLower := Crane.CraneLower;
ActuatorStackVacuumOff := Crane.StackVacuumOff;
ActuatorStackVacuumOn := Crane.StackVacuumOn;
Stamp.StampSliderSensorMovedOut := SensorStampSliderSensorMovedOut;
Stamp.StampSliderSensorMovedIn := SensorStampSliderSensorMovedIn;
Stamp.StampSliderFilled := SensorStampSliderFilled;
Stamp.StampUp := SensorStampUp;
Stamp.StampLowered := SensorStampLowered;
Stamp.CraneDown := SensorCraneDown;
Stamp.CraneUp := SensorCraneUp;
Stamp.CraneSucked := SensorCraneSucked;
Stamp.CranePositionStamp := SensorCranePositionStamp;
Stamp.CraneOnConveyor := SensorCraneOnConveyor;
Stamp.StampStartButton := SensorStampStartButton;
ActuatorStampSliderMovedOut := Stamp.StampSliderMovedOut;
ActuatorStampSliderMovedIn := Stamp.StampSliderMovedIn;
ActuatorStampWhiteLamp := Stamp.StampWhiteLamp;
ActuatorStampPusher := Stamp.StampPusher;
ActuatorStampGreenLamp := Stamp.StampGreenLamp;
ActuatorAnalogCranePressure := 6000;
IF (SensorStampEmergencyStop AND SensorStackEmergencyStop) THEN
    Stack();
    Crane();
    Stamp();
    IF (ActuatorStackGreenLamp AND ActuatorStampGreenLamp) THEN
        IF ((Stamp.StartCommandStamp AND Crane.StartCommandCrane) AND Stack.StartCommandStack) THEN
            Crane.StartVar := TRUE;
            Stack.StartVar := TRUE;
            Stamp.StartVar := TRUE;
        END_IF;
    END_IF;
    Crane.SFCReset := FALSE;
    Stack.SFCReset := FALSE;
    Stamp.SFCReset := FALSE;
ELSIF (NOT SensorStampEmergencyStop OR NOT SensorStackEmergencyStop) THEN
    ActuatorStackSlider := FALSE;
    ActuatorCraneLower := FALSE;
    ActuatorStackVacuumOn := FALSE;
    ActuatorStackVacuumOff := TRUE;
    ActuatorStackGreenLamp := FALSE;
    ActuatorCraneTurnCounterClockwise := FALSE;
    ActuatorCraneTurnClockwise := FALSE;
    ActuatorStampSliderMovedOut := TRUE;
    ActuatorStampSliderMovedIn := FALSE;
    ActuatorStampGreenLamp := FALSE;
    ActuatorStampPusher := FALSE;
    ActuatorAnalogCranePressure := 0;
    Crane.SFCReset := TRUE;
    Stack.SFCReset := TRUE;
    Stamp.SFCReset := TRUE;
    Crane.StartVar := FALSE;
    Stack.StartVar := FALSE;
    Stamp.StartVar := FALSE;
END_IF;
END_PROGRAM

FUNCTION_BLOCK TON
VAR_INPUT
    IN : BOOL;
    PT : TIME;
END_VAR
VAR
    running : BOOL;
END_VAR
VAR_TEMP
    timeout : BOOL;
END_VAR
VAR_OUTPUT
    Q : BOOL;
    ET : TIME;
END_VAR
timeout := NONDETERMINISTIC_BOOL();
IF NOT IN THEN
    Q := FALSE;
    running := FALSE;
ELSIF NOT running AND NOT Q THEN
    running := TRUE;
ELSIF running AND NOT Q THEN
    Q := timeout;
    running := NOT Q;
END_IF;
ET := NONDETERMINISTIC_TIME();
END_FUNCTION_BLOCK
